(* IEC 61131-3 sources: 2026_Projet_YGO_ExcavatriceDragage/TOOLS/TEST_AUTO_CI/RESULTS/H_TREUILS_BENNE/tests (part 4) *)

(* ---- test_fb_winchoutputinterlock.st ---- *)
(* =======================================================================
   🧪 test_fb_winchoutputinterlock.st — FB_WinchOutputInterlock (TC-P10-012, 013, 020, 021, 022, 039.1)
   ───────────────────────────────────────────────────────────────
   Fiche : DOC/AF/AF_Partie-10_Fonction_Winch/FB_WinchOutputInterlock_v1.0.md
   Conventions : 1 appel fb() = 1 scan ; ADVANCE_TIME(10000000) entre les
   scans pour les fronts R_TRIG ; hex décrit en décimal (bit 0 = 1).
   Watchdog frein = 500ms ; RestartDelay = 1500ms ; DeadTimeSameDir/OppositeDir = 1s (défaut).
   Maintien §3bis : DropConfirmDelay = 100ms , MaxSenseHoldTime (T_max) = 1s (défauts, AC8).
   ======================================================================= *)

SETUP
VAR
    fb : FB_WinchOutputInterlock;
END_VAR
END_SETUP

(* ── Remise à zéro commune : Enable=TRUE, frein serré, pause 1500ms pour purger RestartRequired/DeadTime ── *)

TEST 'TC-P10-012 Watchdog frein : BrakeCmd sans confirmation 500ms -> bit0, RestartInhibit, FAULT ; pas de faux defaut au RestartRequired'
    (* Scan 1 : regime nominal, frein serre (BrakeFeedback=FALSE), pause pour purger *)
    fb(Enable := TRUE, Reset := FALSE, SafeStop := FALSE, AscentPermit := TRUE, DescendPermit := TRUE, PowerContactorEngaged := TRUE,
       BrakeFeedback := FALSE, FwdRevSpeedFeedbackOff := TRUE,
       RequestedRelayFwd := FALSE, RequestedRelayRev := FALSE,
       RequestedContactor1 := FALSE, RequestedContactor2 := FALSE,
       RequestedContactor3 := FALSE, RequestedContactor4 := FALSE,
       RequestedStep := 0);
    ADVANCE_TIME(1500000000);
fb(Enable := TRUE, Reset := FALSE, SafeStop := FALSE, AscentPermit := TRUE, DescendPermit := TRUE, PowerContactorEngaged := TRUE,
       BrakeFeedback := FALSE, FwdRevSpeedFeedbackOff := TRUE,
       RequestedRelayFwd := FALSE, RequestedRelayRev := FALSE,
       RequestedContactor1 := FALSE, RequestedContactor2 := FALSE,
       RequestedContactor3 := FALSE, RequestedContactor4 := FALSE,
       RequestedStep := 0);
    ASSERT_TRUE(fb.Ready, 'Regime nominal -> Ready=TRUE');

    (* Scan 2 : demande mouvement, frein NON confirme ouvert (BrakeFeedback=FALSE) -> watchdog arme *)
    ADVANCE_TIME(10000000);
fb(Enable := TRUE, Reset := FALSE, SafeStop := FALSE, AscentPermit := TRUE, DescendPermit := TRUE, PowerContactorEngaged := TRUE,
       BrakeFeedback := FALSE, FwdRevSpeedFeedbackOff := TRUE,
       RequestedRelayFwd := TRUE, RequestedRelayRev := FALSE,
       RequestedContactor1 := TRUE, RequestedContactor2 := FALSE,
       RequestedContactor3 := FALSE, RequestedContactor4 := FALSE,
       RequestedStep := 1);
    ASSERT_TRUE(fb.RelayFwd, 'Demande montee -> RelayFwd');
    ASSERT_TRUE(fb.BrakeCmd, 'Demande montee -> BrakeCmd');
    ASSERT_EQ(fb.State, E_WinchFinalInterlockState.WAIT_BRAKE_COMMAND_CONFIRMATION, 'Etat WAIT_BRAKE_COMMAND_CONFIRMATION (2)');

    (* Scan 3 : apres 500ms sans confirmation -> defaut frein *)
    ADVANCE_TIME(500000000);
fb(Enable := TRUE, Reset := FALSE, SafeStop := FALSE, AscentPermit := TRUE, DescendPermit := TRUE, PowerContactorEngaged := TRUE,
       BrakeFeedback := FALSE, FwdRevSpeedFeedbackOff := TRUE,
       RequestedRelayFwd := TRUE, RequestedRelayRev := FALSE,
       RequestedContactor1 := TRUE, RequestedContactor2 := FALSE,
       RequestedContactor3 := FALSE, RequestedContactor4 := FALSE,
       RequestedStep := 1);
    ASSERT_TRUE(fb.Error, 'Timeout frein 500ms -> Error');
    ASSERT_EQ(fb.ErrorId, 1, 'Timeout frein -> bit0 (1)');
    ASSERT_TRUE(fb.RestartInhibit, 'Timeout frein -> RestartInhibit=TRUE');
    ASSERT_EQ(fb.Reason, E_WinchFinalInterlockReason.BRAKE_COMMAND_NOT_CONFIRMED, 'Reason=BRAKE_COMMAND_NOT_CONFIRMED (1)');
    ASSERT_EQ(fb.State, E_WinchFinalInterlockState.FAULT, 'Etat FAULT (5)');
END_TEST

TEST 'TC-P10-012bis Pas de faux defaut au RestartRequired : BrakeCmd retenu ne doit pas armer le watchdog'
    (* Scan 1 : regime nominal, pause pour purger *)
    fb(Enable := TRUE, Reset := FALSE, SafeStop := FALSE, AscentPermit := TRUE, DescendPermit := TRUE, PowerContactorEngaged := TRUE,
       BrakeFeedback := FALSE, FwdRevSpeedFeedbackOff := TRUE,
       RequestedRelayFwd := FALSE, RequestedRelayRev := FALSE,
       RequestedContactor1 := FALSE, RequestedContactor2 := FALSE,
       RequestedContactor3 := FALSE, RequestedContactor4 := FALSE,
       RequestedStep := 0);
    ADVANCE_TIME(1500000000);
fb(Enable := TRUE, Reset := FALSE, SafeStop := FALSE, AscentPermit := TRUE, DescendPermit := TRUE, PowerContactorEngaged := TRUE,
       BrakeFeedback := FALSE, FwdRevSpeedFeedbackOff := TRUE,
       RequestedRelayFwd := FALSE, RequestedRelayRev := FALSE,
       RequestedContactor1 := FALSE, RequestedContactor2 := FALSE,
       RequestedContactor3 := FALSE, RequestedContactor4 := FALSE,
       RequestedStep := 0);

    (* Scan 2 : demande mouvement, frein confirme (BrakeFeedback=TRUE) -> mouvement autorise *)
    ADVANCE_TIME(10000000);
fb(Enable := TRUE, Reset := FALSE, SafeStop := FALSE, AscentPermit := TRUE, DescendPermit := TRUE, PowerContactorEngaged := TRUE,
       BrakeFeedback := TRUE, FwdRevSpeedFeedbackOff := TRUE,
       RequestedRelayFwd := TRUE, RequestedRelayRev := FALSE,
       RequestedContactor1 := TRUE, RequestedContactor2 := FALSE,
       RequestedContactor3 := FALSE, RequestedContactor4 := FALSE,
       RequestedStep := 1);
    ASSERT_TRUE(fb.RelayFwd, 'Mouvement autorise -> RelayFwd');

    (* Scan 3 : arret -> RestartRequired=TRUE *)
    ADVANCE_TIME(10000000);
fb(Enable := TRUE, Reset := FALSE, SafeStop := FALSE, AscentPermit := TRUE, DescendPermit := TRUE, PowerContactorEngaged := TRUE,
       BrakeFeedback := FALSE, FwdRevSpeedFeedbackOff := TRUE,
       RequestedRelayFwd := FALSE, RequestedRelayRev := FALSE,
       RequestedContactor1 := FALSE, RequestedContactor2 := FALSE,
       RequestedContactor3 := FALSE, RequestedContactor4 := FALSE,
       RequestedStep := 0);

    (* Scan 4 : nouvelle demande IMMEDIATE (RestartRequired=TRUE) -> BrakeCmd retenu, watchdog NON arme *)
    ADVANCE_TIME(10000000);
fb(Enable := TRUE, Reset := FALSE, SafeStop := FALSE, AscentPermit := TRUE, DescendPermit := TRUE, PowerContactorEngaged := TRUE,
       BrakeFeedback := FALSE, FwdRevSpeedFeedbackOff := TRUE,
       RequestedRelayFwd := TRUE, RequestedRelayRev := FALSE,
       RequestedContactor1 := TRUE, RequestedContactor2 := FALSE,
       RequestedContactor3 := FALSE, RequestedContactor4 := FALSE,
       RequestedStep := 1);
    ASSERT_FALSE(fb.RelayFwd, 'RestartRequired -> RelayFwd retenu');
    ASSERT_FALSE(fb.BrakeCmd, 'RestartRequired -> BrakeCmd retenu (FALSE)');
    ASSERT_EQ(fb.State, E_WinchFinalInterlockState.WAIT_RESTART_DELAY, 'Etat WAIT_RESTART_DELAY (4)');

    (* Scan 5 : apres 500ms, BrakeCmd=FALSE -> PAS de faux defaut *)
    ADVANCE_TIME(500000000);
fb(Enable := TRUE, Reset := FALSE, SafeStop := FALSE, AscentPermit := TRUE, DescendPermit := TRUE, PowerContactorEngaged := TRUE,
       BrakeFeedback := FALSE, FwdRevSpeedFeedbackOff := TRUE,
       RequestedRelayFwd := TRUE, RequestedRelayRev := FALSE,
       RequestedContactor1 := TRUE, RequestedContactor2 := FALSE,
       RequestedContactor3 := FALSE, RequestedContactor4 := FALSE,
       RequestedStep := 1);
    ASSERT_FALSE(fb.Error, 'BrakeCmd retenu par RestartRequired -> PAS de faux defaut frein');
    ASSERT_FALSE(fb.RestartInhibit, 'Pas de RestartInhibit sur faux defaut');
END_TEST

TEST 'TC-P10-013 Defaut frein : latches preserves hors Enable, reautorisation complete'
    (* Scan 1 : regime nominal, pause pour purger *)
    fb(Enable := TRUE, Reset := FALSE, SafeStop := FALSE, AscentPermit := TRUE, DescendPermit := TRUE, PowerContactorEngaged := TRUE,
       BrakeFeedback := FALSE, FwdRevSpeedFeedbackOff := TRUE,
       RequestedRelayFwd := FALSE, RequestedRelayRev := FALSE,
       RequestedContactor1 := FALSE, RequestedContactor2 := FALSE,
       RequestedContactor3 := FALSE, RequestedContactor4 := FALSE,
       RequestedStep := 0);
    ADVANCE_TIME(1500000000);
fb(Enable := TRUE, Reset := FALSE, SafeStop := FALSE, AscentPermit := TRUE, DescendPermit := TRUE, PowerContactorEngaged := TRUE,
       BrakeFeedback := FALSE, FwdRevSpeedFeedbackOff := TRUE,
       RequestedRelayFwd := FALSE, RequestedRelayRev := FALSE,
       RequestedContactor1 := FALSE, RequestedContactor2 := FALSE,
       RequestedContactor3 := FALSE, RequestedContactor4 := FALSE,
       RequestedStep := 0);

    (* Scan 2 : demande mouvement, frein non confirme -> watchdog arme *)
    ADVANCE_TIME(10000000);
fb(Enable := TRUE, Reset := FALSE, SafeStop := FALSE, AscentPermit := TRUE, DescendPermit := TRUE, PowerContactorEngaged := TRUE,
       BrakeFeedback := FALSE, FwdRevSpeedFeedbackOff := TRUE,
       RequestedRelayFwd := TRUE, RequestedRelayRev := FALSE,
       RequestedContactor1 := TRUE, RequestedContactor2 := FALSE,
       RequestedContactor3 := FALSE, RequestedContactor4 := FALSE,
       RequestedStep := 1);
    ADVANCE_TIME(500000000);
fb(Enable := TRUE, Reset := FALSE, SafeStop := FALSE, AscentPermit := TRUE, DescendPermit := TRUE, PowerContactorEngaged := TRUE,
       BrakeFeedback := FALSE, FwdRevSpeedFeedbackOff := TRUE,
       RequestedRelayFwd := TRUE, RequestedRelayRev := FALSE,
       RequestedContactor1 := TRUE, RequestedContactor2 := FALSE,
       RequestedContactor3 := FALSE, RequestedContactor4 := FALSE,
       RequestedStep := 1);
    ASSERT_TRUE(fb.Error, 'Precondition : defaut frein');
    ASSERT_TRUE(fb.RestartInhibit, 'Precondition : RestartInhibit');

    (* Scan 3 : Enable=FALSE -> sorties FALSE MAIS latches preserves *)
    ADVANCE_TIME(10000000);
    fb(Enable := FALSE, Reset := FALSE, SafeStop := FALSE, PowerContactorEngaged := TRUE,
       BrakeFeedback := FALSE, FwdRevSpeedFeedbackOff := TRUE,
       RequestedRelayFwd := TRUE, RequestedRelayRev := FALSE,
       RequestedContactor1 := TRUE, RequestedContactor2 := FALSE,
       RequestedContactor3 := FALSE, RequestedContactor4 := FALSE,
       RequestedStep := 1);
    ASSERT_FALSE(fb.RelayFwd, 'Enable=FALSE -> RelayFwd=FALSE');
    ASSERT_FALSE(fb.BrakeCmd, 'Enable=FALSE -> BrakeCmd=FALSE');
    ASSERT_TRUE(fb.RestartInhibit, 'Enable=FALSE -> RestartInhibit PRESERVE');
    ASSERT_EQ(fb.ErrorId, 1, 'Enable=FALSE -> ErrorId bit0 PRESERVE');

    (* Scan 4 : re-Enable, cause disparue (BrakeFeedback=TRUE) + front Reset -> ResetRequired leve *)
    ADVANCE_TIME(10000000);
    fb(Enable := TRUE, Reset := TRUE, SafeStop := FALSE, PowerContactorEngaged := TRUE,
       BrakeFeedback := TRUE, FwdRevSpeedFeedbackOff := TRUE,
       RequestedRelayFwd := FALSE, RequestedRelayRev := FALSE,
       RequestedContactor1 := FALSE, RequestedContactor2 := FALSE,
       RequestedContactor3 := FALSE, RequestedContactor4 := FALSE,
       RequestedStep := 0);
    ADVANCE_TIME(10000000);
fb(Enable := TRUE, Reset := FALSE, SafeStop := FALSE, AscentPermit := TRUE, DescendPermit := TRUE, PowerContactorEngaged := TRUE,
       BrakeFeedback := TRUE, FwdRevSpeedFeedbackOff := TRUE,
       RequestedRelayFwd := FALSE, RequestedRelayRev := FALSE,
       RequestedContactor1 := FALSE, RequestedContactor2 := FALSE,
       RequestedContactor3 := FALSE, RequestedContactor4 := FALSE,
       RequestedStep := 0);
    ASSERT_FALSE(fb.Error, 'Cause disparue + Reset -> Error=FALSE');

    (* Scan 5 : demande neutre observee (MotorRequest=FALSE) -> NeutralRequestSeen *)
    ADVANCE_TIME(10000000);
fb(Enable := TRUE, Reset := FALSE, SafeStop := FALSE, AscentPermit := TRUE, DescendPermit := TRUE, PowerContactorEngaged := TRUE,
       BrakeFeedback := FALSE, FwdRevSpeedFeedbackOff := TRUE,
       RequestedRelayFwd := FALSE, RequestedRelayRev := FALSE,
       RequestedContactor1 := FALSE, RequestedContactor2 := FALSE,
       RequestedContactor3 := FALSE, RequestedContactor4 := FALSE,
       RequestedStep := 0);
    ADVANCE_TIME(1500000000);
fb(Enable := TRUE, Reset := FALSE, SafeStop := FALSE, AscentPermit := TRUE, DescendPermit := TRUE, PowerContactorEngaged := TRUE,
       BrakeFeedback := FALSE, FwdRevSpeedFeedbackOff := TRUE,
       RequestedRelayFwd := FALSE, RequestedRelayRev := FALSE,
       RequestedContactor1 := FALSE, RequestedContactor2 := FALSE,
       RequestedContactor3 := FALSE, RequestedContactor4 := FALSE,
       RequestedStep := 0);

    (* Scan 6 : nouvelle demande distincte -> RestartInhibit leve *)
    ADVANCE_TIME(10000000);
fb(Enable := TRUE, Reset := FALSE, SafeStop := FALSE, AscentPermit := TRUE, DescendPermit := TRUE, PowerContactorEngaged := TRUE,
       BrakeFeedback := TRUE, FwdRevSpeedFeedbackOff := TRUE,
       RequestedRelayFwd := TRUE, RequestedRelayRev := FALSE,
       RequestedContactor1 := TRUE, RequestedContactor2 := FALSE,
       RequestedContactor3 := FALSE, RequestedContactor4 := FALSE,
       RequestedStep := 1);
    ASSERT_FALSE(fb.RestartInhibit, 'Reautorisation complete -> RestartInhibit=FALSE');
    ASSERT_TRUE(fb.RelayFwd, 'Reautorisation -> mouvement autorise');
END_TEST

TEST 'TC-P10-020 Watchdog frein reel terrain : temps/contacteur/bobine'
    (* (essai site — stub) : le watchdog frein reel (temps de reponse contacteur/bobine, usure)
       est une verification terrain sur l automate reel, jamais automatisable en boite noire.
       On verifie ici la brique logicielle : le watchdog 500ms se declenche sur BrakeCmd sans
       confirmation, condition necessaire du diagnostic terrain. *)
    fb(Enable := TRUE, Reset := FALSE, SafeStop := FALSE, AscentPermit := TRUE, DescendPermit := TRUE, PowerContactorEngaged := TRUE,
       BrakeFeedback := FALSE, FwdRevSpeedFeedbackOff := TRUE,
       RequestedRelayFwd := FALSE, RequestedRelayRev := FALSE,
       RequestedContactor1 := FALSE, RequestedContactor2 := FALSE,
       RequestedContactor3 := FALSE, RequestedContactor4 := FALSE,
       RequestedStep := 0);
    ADVANCE_TIME(1500000000);
    // Scan neutre temporise : purge RestartRequired/DeadTimePending (TON tickes apres la pause,
    // comme les ~150 scans de 10ms d'une vraie pause automate) avant la demande mouvement.
fb(Enable := TRUE, Reset := FALSE, SafeStop := FALSE, AscentPermit := TRUE, DescendPermit := TRUE, PowerContactorEngaged := TRUE,
       BrakeFeedback := FALSE, FwdRevSpeedFeedbackOff := TRUE,
       RequestedRelayFwd := FALSE, RequestedRelayRev := FALSE,
       RequestedContactor1 := FALSE, RequestedContactor2 := FALSE,
       RequestedContactor3 := FALSE, RequestedContactor4 := FALSE,
       RequestedStep := 0);
    ADVANCE_TIME(10000000);
fb(Enable := TRUE, Reset := FALSE, SafeStop := FALSE, AscentPermit := TRUE, DescendPermit := TRUE, PowerContactorEngaged := TRUE,
       BrakeFeedback := FALSE, FwdRevSpeedFeedbackOff := TRUE,
       RequestedRelayFwd := TRUE, RequestedRelayRev := FALSE,
       RequestedContactor1 := TRUE, RequestedContactor2 := FALSE,
       RequestedContactor3 := FALSE, RequestedContactor4 := FALSE,
       RequestedStep := 1);
    ADVANCE_TIME(500000000);
fb(Enable := TRUE, Reset := FALSE, SafeStop := FALSE, AscentPermit := TRUE, DescendPermit := TRUE, PowerContactorEngaged := TRUE,
       BrakeFeedback := FALSE, FwdRevSpeedFeedbackOff := TRUE,
       RequestedRelayFwd := TRUE, RequestedRelayRev := FALSE,
       RequestedContactor1 := TRUE, RequestedContactor2 := FALSE,
       RequestedContactor3 := FALSE, RequestedContactor4 := FALSE,
       RequestedStep := 1);
    ASSERT_TRUE(fb.Error, 'Watchdog frein logiciel 500ms -> Error (brique du diagnostic terrain)');
    ASSERT_EQ(fb.Reason, E_WinchFinalInterlockReason.BRAKE_COMMAND_NOT_CONFIRMED, 'Reason=BRAKE_COMMAND_NOT_CONFIRMED');
END_TEST

TEST 'TC-P10-021 Temps mort meme sens : 1s apres arret -> nouvelle demande (DeadTimeSameDir)'
    (* DeadTimeSameDir=2s force pour rendre le temps mort observable (par defaut 1s, masque
       par RestartDelay 1500ms). La demande meme sens est retenue tant que DeadTimeSameDir
       n est pas ecoule. *)
    fb(Enable := TRUE, Reset := FALSE, SafeStop := FALSE, AscentPermit := TRUE, DescendPermit := TRUE, PowerContactorEngaged := TRUE,
       BrakeFeedback := FALSE, FwdRevSpeedFeedbackOff := TRUE,
       RequestedRelayFwd := FALSE, RequestedRelayRev := FALSE,
       RequestedContactor1 := FALSE, RequestedContactor2 := FALSE,
       RequestedContactor3 := FALSE, RequestedContactor4 := FALSE,
       RequestedStep := 0, DeadTimeSameDir := T#2s, DeadTimeOppositeDir := T#2s);
    ADVANCE_TIME(1500000000);
fb(Enable := TRUE, Reset := FALSE, SafeStop := FALSE, AscentPermit := TRUE, DescendPermit := TRUE, PowerContactorEngaged := TRUE,
       BrakeFeedback := FALSE, FwdRevSpeedFeedbackOff := TRUE,
       RequestedRelayFwd := FALSE, RequestedRelayRev := FALSE,
       RequestedContactor1 := FALSE, RequestedContactor2 := FALSE,
       RequestedContactor3 := FALSE, RequestedContactor4 := FALSE,
       RequestedStep := 0, DeadTimeSameDir := T#2s, DeadTimeOppositeDir := T#2s);

    (* Scan 2 : demande montee, frein confirme -> mouvement *)
    ADVANCE_TIME(10000000);
fb(Enable := TRUE, Reset := FALSE, SafeStop := FALSE, AscentPermit := TRUE, DescendPermit := TRUE, PowerContactorEngaged := TRUE,
       BrakeFeedback := TRUE, FwdRevSpeedFeedbackOff := TRUE,
       RequestedRelayFwd := TRUE, RequestedRelayRev := FALSE,
       RequestedContactor1 := TRUE, RequestedContactor2 := FALSE,
       RequestedContactor3 := FALSE, RequestedContactor4 := FALSE,
       RequestedStep := 1, DeadTimeSameDir := T#2s, DeadTimeOppositeDir := T#2s);
    ASSERT_TRUE(fb.RelayFwd, 'Mouvement autorise -> RelayFwd');

    (* Scan 3 : arret -> DeadTimePending=TRUE *)
    ADVANCE_TIME(10000000);
fb(Enable := TRUE, Reset := FALSE, SafeStop := FALSE, AscentPermit := TRUE, DescendPermit := TRUE, PowerContactorEngaged := TRUE,
       BrakeFeedback := FALSE, FwdRevSpeedFeedbackOff := TRUE,
       RequestedRelayFwd := FALSE, RequestedRelayRev := FALSE,
       RequestedContactor1 := FALSE, RequestedContactor2 := FALSE,
       RequestedContactor3 := FALSE, RequestedContactor4 := FALSE,
       RequestedStep := 0, DeadTimeSameDir := T#2s, DeadTimeOppositeDir := T#2s);

    (* Scan 4 : apres 1500ms (RestartRequired leve), DeadTimeSameDir=2s pas encore ecoule -> retenu *)
    ADVANCE_TIME(1500000000);
fb(Enable := TRUE, Reset := FALSE, SafeStop := FALSE, AscentPermit := TRUE, DescendPermit := TRUE, PowerContactorEngaged := TRUE,
       BrakeFeedback := FALSE, FwdRevSpeedFeedbackOff := TRUE,
       RequestedRelayFwd := TRUE, RequestedRelayRev := FALSE,
       RequestedContactor1 := TRUE, RequestedContactor2 := FALSE,
       RequestedContactor3 := FALSE, RequestedContactor4 := FALSE,
       RequestedStep := 1, DeadTimeSameDir := T#2s, DeadTimeOppositeDir := T#2s);
    ASSERT_FALSE(fb.RelayFwd, 'DeadTimeSameDir pas ecoule -> demande meme sens retenue');
    ASSERT_EQ(fb.State, E_WinchFinalInterlockState.WAIT_RESTART_DELAY, 'Etat WAIT_RESTART_DELAY (4)');

    (* Scan 5 : apres 2s (DeadTimeSameDir ecoule) -> demande meme sens acceptee *)
    ADVANCE_TIME(600000000);
fb(Enable := TRUE, Reset := FALSE, SafeStop := FALSE, AscentPermit := TRUE, DescendPermit := TRUE, PowerContactorEngaged := TRUE,
       BrakeFeedback := TRUE, FwdRevSpeedFeedbackOff := TRUE,
       RequestedRelayFwd := TRUE, RequestedRelayRev := FALSE,
       RequestedContactor1 := TRUE, RequestedContactor2 := FALSE,
       RequestedContactor3 := FALSE, RequestedContactor4 := FALSE,
       RequestedStep := 1, DeadTimeSameDir := T#2s, DeadTimeOppositeDir := T#2s);
    ASSERT_TRUE(fb.RelayFwd, 'DeadTimeSameDir ecoule -> demande meme sens acceptee');
END_TEST

TEST 'TC-P10-022 Temps mort inversion : 1s apres arret + inversion sens (DeadTimeOppositeDir)'
    (* DeadTimeOppositeDir=2s force pour rendre le temps mort d inversion observable.
       L inversion est retenue tant que DeadTimeOppositeDir n est pas ecoule. *)
    fb(Enable := TRUE, Reset := FALSE, SafeStop := FALSE, AscentPermit := TRUE, DescendPermit := TRUE, PowerContactorEngaged := TRUE,
       BrakeFeedback := FALSE, FwdRevSpeedFeedbackOff := TRUE,
       RequestedRelayFwd := FALSE, RequestedRelayRev := FALSE,
       RequestedContactor1 := FALSE, RequestedContactor2 := FALSE,
       RequestedContactor3 := FALSE, RequestedContactor4 := FALSE,
       RequestedStep := 0, DeadTimeSameDir := T#1s, DeadTimeOppositeDir := T#2s);
    ADVANCE_TIME(1500000000);
fb(Enable := TRUE, Reset := FALSE, SafeStop := FALSE, AscentPermit := TRUE, DescendPermit := TRUE, PowerContactorEngaged := TRUE,
       BrakeFeedback := FALSE, FwdRevSpeedFeedbackOff := TRUE,
       RequestedRelayFwd := FALSE, RequestedRelayRev := FALSE,
       RequestedContactor1 := FALSE, RequestedContactor2 := FALSE,
       RequestedContactor3 := FALSE, RequestedContactor4 := FALSE,
       RequestedStep := 0, DeadTimeSameDir := T#1s, DeadTimeOppositeDir := T#2s);

    (* Scan 2 : demande montee, frein confirme -> mouvement *)
    ADVANCE_TIME(10000000);
fb(Enable := TRUE, Reset := FALSE, SafeStop := FALSE, AscentPermit := TRUE, DescendPermit := TRUE, PowerContactorEngaged := TRUE,
       BrakeFeedback := TRUE, FwdRevSpeedFeedbackOff := TRUE,
       RequestedRelayFwd := TRUE, RequestedRelayRev := FALSE,
       RequestedContactor1 := TRUE, RequestedContactor2 := FALSE,
       RequestedContactor3 := FALSE, RequestedContactor4 := FALSE,
       RequestedStep := 1, DeadTimeSameDir := T#1s, DeadTimeOppositeDir := T#2s);
    ASSERT_TRUE(fb.RelayFwd, 'Mouvement montee -> RelayFwd');

    (* Scan 3 : arret -> DeadTimePending=TRUE *)
    ADVANCE_TIME(10000000);
fb(Enable := TRUE, Reset := FALSE, SafeStop := FALSE, AscentPermit := TRUE, DescendPermit := TRUE, PowerContactorEngaged := TRUE,
       BrakeFeedback := FALSE, FwdRevSpeedFeedbackOff := TRUE,
       RequestedRelayFwd := FALSE, RequestedRelayRev := FALSE,
       RequestedContactor1 := FALSE, RequestedContactor2 := FALSE,
       RequestedContactor3 := FALSE, RequestedContactor4 := FALSE,
       RequestedStep := 0, DeadTimeSameDir := T#1s, DeadTimeOppositeDir := T#2s);

    (* Scan 4 : apres 1500ms, inversion (descente) -> DeadTimeOppositeDir=2s pas ecoule -> retenu *)
    ADVANCE_TIME(1500000000);
fb(Enable := TRUE, Reset := FALSE, SafeStop := FALSE, AscentPermit := TRUE, DescendPermit := TRUE, PowerContactorEngaged := TRUE,
       BrakeFeedback := FALSE, FwdRevSpeedFeedbackOff := TRUE,
       RequestedRelayFwd := FALSE, RequestedRelayRev := TRUE,
       RequestedContactor1 := TRUE, RequestedContactor2 := FALSE,
       RequestedContactor3 := FALSE, RequestedContactor4 := FALSE,
       RequestedStep := 1, DeadTimeSameDir := T#1s, DeadTimeOppositeDir := T#2s);
    ASSERT_FALSE(fb.RelayRev, 'DeadTimeOppositeDir pas ecoule -> inversion retenue');
    ASSERT_EQ(fb.State, E_WinchFinalInterlockState.WAIT_RESTART_DELAY, 'Etat WAIT_RESTART_DELAY (4)');

    (* Scan 5 : apres 2s (DeadTimeOppositeDir ecoule) -> inversion acceptee *)
    ADVANCE_TIME(600000000);
fb(Enable := TRUE, Reset := FALSE, SafeStop := FALSE, AscentPermit := TRUE, DescendPermit := TRUE, PowerContactorEngaged := TRUE,
       BrakeFeedback := TRUE, FwdRevSpeedFeedbackOff := TRUE,
       RequestedRelayFwd := FALSE, RequestedRelayRev := TRUE,
       RequestedContactor1 := TRUE, RequestedContactor2 := FALSE,
       RequestedContactor3 := FALSE, RequestedContactor4 := FALSE,
       RequestedStep := 1, DeadTimeSameDir := T#1s, DeadTimeOppositeDir := T#2s);
    ASSERT_TRUE(fb.RelayRev, 'DeadTimeOppositeDir ecoule -> inversion acceptee');
END_TEST

TEST 'TC-P10-039.1 Frein couple direct : BrakeCmd = RelayFwd OR RelayRev dans tous les etats'
    (* Scan 1 : regime nominal, pause pour purger *)
    fb(Enable := TRUE, Reset := FALSE, SafeStop := FALSE, AscentPermit := TRUE, DescendPermit := TRUE, PowerContactorEngaged := TRUE,
       BrakeFeedback := FALSE, FwdRevSpeedFeedbackOff := TRUE,
       RequestedRelayFwd := FALSE, RequestedRelayRev := FALSE,
       RequestedContactor1 := FALSE, RequestedContactor2 := FALSE,
       RequestedContactor3 := FALSE, RequestedContactor4 := FALSE,
       RequestedStep := 0);
    ADVANCE_TIME(1500000000);
fb(Enable := TRUE, Reset := FALSE, SafeStop := FALSE, AscentPermit := TRUE, DescendPermit := TRUE, PowerContactorEngaged := TRUE,
       BrakeFeedback := FALSE, FwdRevSpeedFeedbackOff := TRUE,
       RequestedRelayFwd := FALSE, RequestedRelayRev := FALSE,
       RequestedContactor1 := FALSE, RequestedContactor2 := FALSE,
       RequestedContactor3 := FALSE, RequestedContactor4 := FALSE,
       RequestedStep := 0);
    ASSERT_FALSE(fb.BrakeCmd, 'Repos : BrakeCmd=FALSE (RelayFwd/Rev=FALSE)');

    (* Scan 2 : mouvement montee -> BrakeCmd=TRUE (RelayFwd=TRUE) *)
    ADVANCE_TIME(10000000);
fb(Enable := TRUE, Reset := FALSE, SafeStop := FALSE, AscentPermit := TRUE, DescendPermit := TRUE, PowerContactorEngaged := TRUE,
       BrakeFeedback := TRUE, FwdRevSpeedFeedbackOff := TRUE,
       RequestedRelayFwd := TRUE, RequestedRelayRev := FALSE,
       RequestedContactor1 := TRUE, RequestedContactor2 := FALSE,
       RequestedContactor3 := FALSE, RequestedContactor4 := FALSE,
       RequestedStep := 1);
    ASSERT_TRUE(fb.RelayFwd, 'Mouvement -> RelayFwd=TRUE');
    ASSERT_TRUE(fb.BrakeCmd, 'Mouvement -> BrakeCmd=TRUE (couple direct)');

    (* Scan 3 : arret -> BrakeCmd=FALSE *)
    ADVANCE_TIME(10000000);
fb(Enable := TRUE, Reset := FALSE, SafeStop := FALSE, AscentPermit := TRUE, DescendPermit := TRUE, PowerContactorEngaged := TRUE,
       BrakeFeedback := FALSE, FwdRevSpeedFeedbackOff := TRUE,
       RequestedRelayFwd := FALSE, RequestedRelayRev := FALSE,
       RequestedContactor1 := FALSE, RequestedContactor2 := FALSE,
       RequestedContactor3 := FALSE, RequestedContactor4 := FALSE,
       RequestedStep := 0);
    ASSERT_FALSE(fb.RelayFwd, 'Arret -> RelayFwd=FALSE');
    ASSERT_FALSE(fb.BrakeCmd, 'Arret -> BrakeCmd=FALSE (jamais de divergence frein/mouvement)');
END_TEST

TEST 'TC-P10-023a §3bis : sens maintenu apres chute de palier a 0 tant que contacteurs non confirmes, puis chute sur DropConfirmDelay'
    (* Chute de palier : RequestedStep -> 0 mais RequestedRelayFwd reste TRUE (demande transitoire
       FB_Winch). La barriere TIENT le contacteur de sens jusqu a FwdRevSpeedFeedbackOff confirme
       (debounced DropConfirmDelay=300ms) OU T_max. Aucun faux arret pendant le debounce. *)
    fb(Enable := TRUE, Reset := FALSE, SafeStop := FALSE, AscentPermit := TRUE, DescendPermit := TRUE, PowerContactorEngaged := TRUE,
       BrakeFeedback := FALSE, FwdRevSpeedFeedbackOff := TRUE,
       RequestedRelayFwd := FALSE, RequestedRelayRev := FALSE,
       RequestedContactor1 := FALSE, RequestedContactor2 := FALSE,
       RequestedContactor3 := FALSE, RequestedContactor4 := FALSE,
       RequestedStep := 0, DropConfirmDelay := T#300ms, MaxSenseHoldTime := T#1s);
    ADVANCE_TIME(1500000000);
fb(Enable := TRUE, Reset := FALSE, SafeStop := FALSE, AscentPermit := TRUE, DescendPermit := TRUE, PowerContactorEngaged := TRUE,
       BrakeFeedback := FALSE, FwdRevSpeedFeedbackOff := TRUE,
       RequestedRelayFwd := FALSE, RequestedRelayRev := FALSE,
       RequestedContactor1 := FALSE, RequestedContactor2 := FALSE,
       RequestedContactor3 := FALSE, RequestedContactor4 := FALSE,
       RequestedStep := 0, DropConfirmDelay := T#300ms, MaxSenseHoldTime := T#1s);
    ASSERT_TRUE(fb.Ready, 'Regime nominal -> Ready=TRUE');

    (* Scan 2 : mouvement montee, frein confirme, contacteurs engages (FwdRevSpeedFeedbackOff=FALSE) *)
    ADVANCE_TIME(10000000);
fb(Enable := TRUE, Reset := FALSE, SafeStop := FALSE, AscentPermit := TRUE, DescendPermit := TRUE, PowerContactorEngaged := TRUE,
       BrakeFeedback := TRUE, FwdRevSpeedFeedbackOff := FALSE,
       RequestedRelayFwd := TRUE, RequestedRelayRev := FALSE,
       RequestedContactor1 := TRUE, RequestedContactor2 := FALSE,
       RequestedContactor3 := FALSE, RequestedContactor4 := FALSE,
       RequestedStep := 1, DropConfirmDelay := T#300ms, MaxSenseHoldTime := T#1s);
    ASSERT_TRUE(fb.RelayFwd, 'Mouvement -> RelayFwd');
    ASSERT_TRUE(fb.BrakeCmd, 'Mouvement -> BrakeCmd');

    (* Scan 3 : chute a palier 0, RequestedRelayFwd TOUJOURS TRUE, contacteurs pas encore retombes *)
    ADVANCE_TIME(10000000);
fb(Enable := TRUE, Reset := FALSE, SafeStop := FALSE, AscentPermit := TRUE, DescendPermit := TRUE, PowerContactorEngaged := TRUE,
       BrakeFeedback := TRUE, FwdRevSpeedFeedbackOff := FALSE,
       RequestedRelayFwd := TRUE, RequestedRelayRev := FALSE,
       RequestedContactor1 := FALSE, RequestedContactor2 := FALSE,
       RequestedContactor3 := FALSE, RequestedContactor4 := FALSE,
       RequestedStep := 0, DropConfirmDelay := T#300ms, MaxSenseHoldTime := T#1s);
    ASSERT_TRUE(fb.RelayFwd, 'Chute palier -> contacteur de sens MAINTENU (§3bis)');
    ASSERT_TRUE(fb.BrakeCmd, 'Maintien -> BrakeCmd reste TRUE (couple direct)');
    ASSERT_TRUE(fb.SenseHoldActive, 'Diag SenseHoldActive');
    ASSERT_EQ(fb.State, E_WinchFinalInterlockState.WAIT_SENSE_DROP_CONFIRM, 'Etat WAIT_SENSE_DROP_CONFIRM (6)');

    (* Scan 4 : feedback retombee percu (FwdRevSpeedFeedbackOff=TRUE) mais debounce pas ecoule -> tenu *)
    ADVANCE_TIME(100000000);
fb(Enable := TRUE, Reset := FALSE, SafeStop := FALSE, AscentPermit := TRUE, DescendPermit := TRUE, PowerContactorEngaged := TRUE,
       BrakeFeedback := TRUE, FwdRevSpeedFeedbackOff := TRUE,
       RequestedRelayFwd := TRUE, RequestedRelayRev := FALSE,
       RequestedContactor1 := FALSE, RequestedContactor2 := FALSE,
       RequestedContactor3 := FALSE, RequestedContactor4 := FALSE,
       RequestedStep := 0, DropConfirmDelay := T#300ms, MaxSenseHoldTime := T#1s);
    ASSERT_TRUE(fb.RelayFwd, 'Debounce DropConfirmDelay pas ecoule -> sens TOUJOURS tenu (AC7)');

    (* Scan 5 : DropConfirmDelay (300ms) ecoule -> chute normale du sens *)
    ADVANCE_TIME(300000000);
fb(Enable := TRUE, Reset := FALSE, SafeStop := FALSE, AscentPermit := TRUE, DescendPermit := TRUE, PowerContactorEngaged := TRUE,
       BrakeFeedback := TRUE, FwdRevSpeedFeedbackOff := TRUE,
       RequestedRelayFwd := TRUE, RequestedRelayRev := FALSE,
       RequestedContactor1 := FALSE, RequestedContactor2 := FALSE,
       RequestedContactor3 := FALSE, RequestedContactor4 := FALSE,
       RequestedStep := 0, DropConfirmDelay := T#300ms, MaxSenseHoldTime := T#1s);
    ADVANCE_TIME(10000000);
fb(Enable := TRUE, Reset := FALSE, SafeStop := FALSE, AscentPermit := TRUE, DescendPermit := TRUE, PowerContactorEngaged := TRUE,
       BrakeFeedback := TRUE, FwdRevSpeedFeedbackOff := TRUE,
       RequestedRelayFwd := TRUE, RequestedRelayRev := FALSE,
       RequestedContactor1 := FALSE, RequestedContactor2 := FALSE,
       RequestedContactor3 := FALSE, RequestedContactor4 := FALSE,
       RequestedStep := 0, DropConfirmDelay := T#300ms, MaxSenseHoldTime := T#1s);
    ASSERT_FALSE(fb.RelayFwd, 'Confirmation retombee -> chute du sens (§3bis)');
    ASSERT_FALSE(fb.BrakeCmd, 'Apres chute -> BrakeCmd=FALSE');
    ASSERT_FALSE(fb.SenseHoldActive, 'Fin du maintien');
    ASSERT_EQ(fb.State, E_WinchFinalInterlockState.READY, 'Retour READY');
END_TEST

TEST 'TC-P10-023b §3bis : T_max atteint sans confirmation -> chute du sens FORCEE + latch ContactorStuck'
    (* FwdRevSpeedFeedbackOff reste FALSE (contacteurs ne confirment pas la retombee). Apres
       MaxSenseHoldTime (T_max=300ms) la barriere FORCE la chute du sens et latche
       ContactorStuck (AC7). Le maintien indefini du stator est interdit. *)
    fb(Enable := TRUE, Reset := FALSE, SafeStop := FALSE, AscentPermit := TRUE, DescendPermit := TRUE, PowerContactorEngaged := TRUE,
       BrakeFeedback := FALSE, FwdRevSpeedFeedbackOff := TRUE,
       RequestedRelayFwd := FALSE, RequestedRelayRev := FALSE,
       RequestedContactor1 := FALSE, RequestedContactor2 := FALSE,
       RequestedContactor3 := FALSE, RequestedContactor4 := FALSE,
       RequestedStep := 0, DropConfirmDelay := T#200ms, MaxSenseHoldTime := T#300ms);
    ADVANCE_TIME(1500000000);
fb(Enable := TRUE, Reset := FALSE, SafeStop := FALSE, AscentPermit := TRUE, DescendPermit := TRUE, PowerContactorEngaged := TRUE,
       BrakeFeedback := FALSE, FwdRevSpeedFeedbackOff := TRUE,
       RequestedRelayFwd := FALSE, RequestedRelayRev := FALSE,
       RequestedContactor1 := FALSE, RequestedContactor2 := FALSE,
       RequestedContactor3 := FALSE, RequestedContactor4 := FALSE,
       RequestedStep := 0, DropConfirmDelay := T#200ms, MaxSenseHoldTime := T#300ms);

    (* Scan 2 : mouvement montee *)
    ADVANCE_TIME(10000000);
fb(Enable := TRUE, Reset := FALSE, SafeStop := FALSE, AscentPermit := TRUE, DescendPermit := TRUE, PowerContactorEngaged := TRUE,
       BrakeFeedback := TRUE, FwdRevSpeedFeedbackOff := FALSE,
       RequestedRelayFwd := TRUE, RequestedRelayRev := FALSE,
       RequestedContactor1 := TRUE, RequestedContactor2 := FALSE,
       RequestedContactor3 := FALSE, RequestedContactor4 := FALSE,
       RequestedStep := 1, DropConfirmDelay := T#200ms, MaxSenseHoldTime := T#300ms);
    ASSERT_TRUE(fb.RelayFwd, 'Mouvement -> RelayFwd');

    (* Scan 3 : chute palier a 0, sens maintenu, MAIS contacteurs jamais confirmes retombes *)
    ADVANCE_TIME(10000000);
fb(Enable := TRUE, Reset := FALSE, SafeStop := FALSE, AscentPermit := TRUE, DescendPermit := TRUE, PowerContactorEngaged := TRUE,
       BrakeFeedback := TRUE, FwdRevSpeedFeedbackOff := FALSE,
       RequestedRelayFwd := TRUE, RequestedRelayRev := FALSE,
       RequestedContactor1 := FALSE, RequestedContactor2 := FALSE,
       RequestedContactor3 := FALSE, RequestedContactor4 := FALSE,
       RequestedStep := 0, DropConfirmDelay := T#200ms, MaxSenseHoldTime := T#300ms);
    ASSERT_TRUE(fb.RelayFwd, 'Entree en maintien -> sens tenu');
    ASSERT_TRUE(fb.SenseHoldActive, 'SenseHoldActive');

    (* Scan 4 : T_max (300ms) depasse sans confirmation -> chute forcee + latch *)
    ADVANCE_TIME(10000000);
fb(Enable := TRUE, Reset := FALSE, SafeStop := FALSE, AscentPermit := TRUE, DescendPermit := TRUE, PowerContactorEngaged := TRUE,
       BrakeFeedback := TRUE, FwdRevSpeedFeedbackOff := FALSE,
       RequestedRelayFwd := TRUE, RequestedRelayRev := FALSE,
       RequestedContactor1 := FALSE, RequestedContactor2 := FALSE,
       RequestedContactor3 := FALSE, RequestedContactor4 := FALSE,
       RequestedStep := 0, DropConfirmDelay := T#200ms, MaxSenseHoldTime := T#300ms);
    ADVANCE_TIME(400000000);
fb(Enable := TRUE, Reset := FALSE, SafeStop := FALSE, AscentPermit := TRUE, DescendPermit := TRUE, PowerContactorEngaged := TRUE,
       BrakeFeedback := TRUE, FwdRevSpeedFeedbackOff := FALSE,
       RequestedRelayFwd := TRUE, RequestedRelayRev := FALSE,
       RequestedContactor1 := FALSE, RequestedContactor2 := FALSE,
       RequestedContactor3 := FALSE, RequestedContactor4 := FALSE,
       RequestedStep := 0, DropConfirmDelay := T#200ms, MaxSenseHoldTime := T#300ms);
    ASSERT_FALSE(fb.RelayFwd, 'T_max sans confirmation -> chute du sens FORCEE (AC7)');
    ASSERT_FALSE(fb.BrakeCmd, 'Chute forcee -> BrakeCmd=FALSE');
    ASSERT_TRUE(fb.ContactorStuck, 'Diag ContactorStuck latche');
    ASSERT_FALSE(fb.SenseHoldActive, 'Fin du maintien');
    ASSERT_FALSE(fb.Ready, 'Latch -> barriere non pret (pas de redemarrage auto)');
    ASSERT_EQ(fb.State, E_WinchFinalInterlockState.FAULT, 'Etat FAULT');
    ASSERT_EQ(fb.Reason, E_WinchFinalInterlockReason.SENSE_DROP_TIMEOUT, 'Reason=SENSE_DROP_TIMEOUT');

    (* Scan 5 : acquittement conscient (front Reset) -> latch leve (cause disparue = demande neutre) *)
    ADVANCE_TIME(10000000);
    fb(Enable := TRUE, Reset := TRUE, SafeStop := FALSE, PowerContactorEngaged := TRUE,
       BrakeFeedback := TRUE, FwdRevSpeedFeedbackOff := TRUE,
       RequestedRelayFwd := FALSE, RequestedRelayRev := FALSE,
       RequestedContactor1 := FALSE, RequestedContactor2 := FALSE,
       RequestedContactor3 := FALSE, RequestedContactor4 := FALSE,
       RequestedStep := 0, DropConfirmDelay := T#200ms, MaxSenseHoldTime := T#300ms);
    ADVANCE_TIME(10000000);
fb(Enable := TRUE, Reset := FALSE, SafeStop := FALSE, AscentPermit := TRUE, DescendPermit := TRUE, PowerContactorEngaged := TRUE,
       BrakeFeedback := TRUE, FwdRevSpeedFeedbackOff := TRUE,
       RequestedRelayFwd := FALSE, RequestedRelayRev := FALSE,
       RequestedContactor1 := FALSE, RequestedContactor2 := FALSE,
       RequestedContactor3 := FALSE, RequestedContactor4 := FALSE,
       RequestedStep := 0, DropConfirmDelay := T#200ms, MaxSenseHoldTime := T#300ms);
    ASSERT_FALSE(fb.ContactorStuck, 'Front Reset conscient -> latch ContactorStuck leve');
END_TEST

TEST 'TC-P10-023c §3bis : coupure dure (Enable=FALSE) pendant le maintien -> RelayFwd=FALSE immediat'
    (* La coupure dure ne passe JAMAIS par le maintien §3bis (AC9) : Enable=FALSE en pleine
       tenue du sens coupe RelayFwd/Rev au cycle suivant, sans attendre confirmation ni T_max. *)
    fb(Enable := TRUE, Reset := FALSE, SafeStop := FALSE, AscentPermit := TRUE, DescendPermit := TRUE, PowerContactorEngaged := TRUE,
       BrakeFeedback := FALSE, FwdRevSpeedFeedbackOff := TRUE,
       RequestedRelayFwd := FALSE, RequestedRelayRev := FALSE,
       RequestedContactor1 := FALSE, RequestedContactor2 := FALSE,
       RequestedContactor3 := FALSE, RequestedContactor4 := FALSE,
       RequestedStep := 0, DropConfirmDelay := T#300ms, MaxSenseHoldTime := T#1s);
    ADVANCE_TIME(1500000000);
fb(Enable := TRUE, Reset := FALSE, SafeStop := FALSE, AscentPermit := TRUE, DescendPermit := TRUE, PowerContactorEngaged := TRUE,
       BrakeFeedback := FALSE, FwdRevSpeedFeedbackOff := TRUE,
       RequestedRelayFwd := FALSE, RequestedRelayRev := FALSE,
       RequestedContactor1 := FALSE, RequestedContactor2 := FALSE,
       RequestedContactor3 := FALSE, RequestedContactor4 := FALSE,
       RequestedStep := 0, DropConfirmDelay := T#300ms, MaxSenseHoldTime := T#1s);

    (* Scan 2 : mouvement montee *)
    ADVANCE_TIME(10000000);
fb(Enable := TRUE, Reset := FALSE, SafeStop := FALSE, AscentPermit := TRUE, DescendPermit := TRUE, PowerContactorEngaged := TRUE,
       BrakeFeedback := TRUE, FwdRevSpeedFeedbackOff := FALSE,
       RequestedRelayFwd := TRUE, RequestedRelayRev := FALSE,
       RequestedContactor1 := TRUE, RequestedContactor2 := FALSE,
       RequestedContactor3 := FALSE, RequestedContactor4 := FALSE,
       RequestedStep := 1, DropConfirmDelay := T#300ms, MaxSenseHoldTime := T#1s);
    ASSERT_TRUE(fb.RelayFwd, 'Mouvement -> RelayFwd');

    (* Scan 3 : chute palier a 0 -> maintien actif *)
    ADVANCE_TIME(10000000);
fb(Enable := TRUE, Reset := FALSE, SafeStop := FALSE, AscentPermit := TRUE, DescendPermit := TRUE, PowerContactorEngaged := TRUE,
       BrakeFeedback := TRUE, FwdRevSpeedFeedbackOff := FALSE,
       RequestedRelayFwd := TRUE, RequestedRelayRev := FALSE,
       RequestedContactor1 := FALSE, RequestedContactor2 := FALSE,
       RequestedContactor3 := FALSE, RequestedContactor4 := FALSE,
       RequestedStep := 0, DropConfirmDelay := T#300ms, MaxSenseHoldTime := T#1s);
    ASSERT_TRUE(fb.RelayFwd, 'Maintien actif -> sens tenu');
    ASSERT_TRUE(fb.SenseHoldActive, 'SenseHoldActive');

    (* Scan 4 : Enable=FALSE -> coupure dure immediate, meme en pleine tenue *)
    ADVANCE_TIME(10000000);
    fb(Enable := FALSE, Reset := FALSE, SafeStop := FALSE, PowerContactorEngaged := TRUE,
       BrakeFeedback := TRUE, FwdRevSpeedFeedbackOff := FALSE,
       RequestedRelayFwd := TRUE, RequestedRelayRev := FALSE,
       RequestedContactor1 := FALSE, RequestedContactor2 := FALSE,
       RequestedContactor3 := FALSE, RequestedContactor4 := FALSE,
       RequestedStep := 0, DropConfirmDelay := T#300ms, MaxSenseHoldTime := T#1s);
    ASSERT_FALSE(fb.RelayFwd, 'Enable=FALSE -> RelayFwd=FALSE immediat (AC9)');
    ASSERT_FALSE(fb.BrakeCmd, 'Enable=FALSE -> BrakeCmd=FALSE immediat');
    ASSERT_FALSE(fb.SenseHoldActive, 'Maintien neutralise par la gate');
END_TEST

TEST 'TC-T216-FINAL-PERMIT Direction refusee coupe la barriere finale, direction autorisee passe'
    (* Le permis final est une defense en profondeur : il doit couper relais,
       contacteurs et frein meme si une demande physique est encore presente. *)
    fb(Enable := TRUE, Reset := FALSE, SafeStop := FALSE, AscentPermit := TRUE, DescendPermit := TRUE,
       PowerContactorEngaged := TRUE, BrakeFeedback := TRUE, FwdRevSpeedFeedbackOff := TRUE,
       RequestedRelayFwd := TRUE, RequestedRelayRev := FALSE,
       RequestedContactor1 := TRUE, RequestedContactor2 := FALSE,
       RequestedContactor3 := FALSE, RequestedContactor4 := FALSE, RequestedStep := 1);
    ASSERT_TRUE(fb.RelayFwd, 'Permis montee TRUE -> relais montee autorise');
    ASSERT_TRUE(fb.BrakeCmd, 'Permis montee TRUE -> frein desserre');

    ADVANCE_TIME(10000000);
    fb(Enable := TRUE, Reset := FALSE, SafeStop := FALSE, AscentPermit := FALSE, DescendPermit := TRUE,
       PowerContactorEngaged := TRUE, BrakeFeedback := TRUE, FwdRevSpeedFeedbackOff := TRUE,
       RequestedRelayFwd := TRUE, RequestedRelayRev := FALSE,
       RequestedContactor1 := TRUE, RequestedContactor2 := FALSE,
       RequestedContactor3 := FALSE, RequestedContactor4 := FALSE, RequestedStep := 1);
    ASSERT_FALSE(fb.RelayFwd, 'Permis montee FALSE -> relais montee coupe');
    ASSERT_FALSE(fb.Contactor1, 'Permis montee FALSE -> contacteur coupe');
    ASSERT_FALSE(fb.BrakeCmd, 'Permis montee FALSE -> frein serre');

    ADVANCE_TIME(10000000);
    fb(Enable := TRUE, Reset := FALSE, SafeStop := FALSE, AscentPermit := TRUE, DescendPermit := FALSE,
       PowerContactorEngaged := TRUE, BrakeFeedback := TRUE, FwdRevSpeedFeedbackOff := TRUE,
       RequestedRelayFwd := FALSE, RequestedRelayRev := TRUE,
       RequestedContactor1 := TRUE, RequestedContactor2 := FALSE,
       RequestedContactor3 := FALSE, RequestedContactor4 := FALSE, RequestedStep := 1);
    ASSERT_FALSE(fb.RelayRev, 'Permis descente FALSE -> relais descente coupe');
    ASSERT_FALSE(fb.Contactor1, 'Permis descente FALSE -> contacteur coupe');
    ASSERT_FALSE(fb.BrakeCmd, 'Permis descente FALSE -> frein serre');
END_TEST

(* ---- test_fb_winchstepshaper.st ---- *)
SETUP
VAR
    fb : FB_WinchStepShaper;
END_VAR
END_SETUP

TEST 'TC-P10-SHAPER-01 Montee nominale 1000ms'
    fb(Enable := TRUE, TargetStep := 0, StepRampDelay := T#1000ms);
    ASSERT_EQ(fb.ShapedStep, 0, 'ShapedStep initialement a 0');

    (* Depart immediat 0->1 au scan 0 *)
    fb(Enable := TRUE, TargetStep := 5, StepRampDelay := T#1000ms);
    ASSERT_EQ(fb.ShapedStep, 1, 'ShapedStep passe a 1 immediatement');

    (* Echantillonnage avant delai *)
    ADVANCE_TIME(10000000);
    fb(Enable := TRUE, TargetStep := 5, StepRampDelay := T#1000ms);
    ASSERT_EQ(fb.ShapedStep, 1, 'Reste a 1 avant delai');

    (* Ecoulement 1000ms -> P2 *)
    ADVANCE_TIME(1000000000);
    fb(Enable := TRUE, TargetStep := 5, StepRampDelay := T#1000ms);
    ASSERT_EQ(fb.ShapedStep, 2, 'Passe a 2 apres delai');
END_TEST

TEST 'TC-P10-SHAPER-02 Descente nominale 500ms'
    fb(Enable := TRUE, TargetStep := 2, StepRampDelay := T#500ms);
    ASSERT_EQ(fb.ShapedStep, 1, 'Depart P1');

    ADVANCE_TIME(10000000);
    fb(Enable := TRUE, TargetStep := 2, StepRampDelay := T#500ms);
    ASSERT_EQ(fb.ShapedStep, 1, 'Reste a 1');

    ADVANCE_TIME(500000000);
    fb(Enable := TRUE, TargetStep := 2, StepRampDelay := T#500ms);
    ASSERT_EQ(fb.ShapedStep, 2, 'Passe a 2 apres delai 500ms');
END_TEST

TEST 'TC-P10-SHAPER-03 Asymetrie arret direct'
    fb(Enable := TRUE, TargetStep := 2, StepRampDelay := T#500ms);
    ASSERT_EQ(fb.ShapedStep, 1, 'Depart P1');

    ADVANCE_TIME(10000000);
    fb(Enable := TRUE, TargetStep := 2, StepRampDelay := T#500ms);
    ADVANCE_TIME(500000000);
    fb(Enable := TRUE, TargetStep := 2, StepRampDelay := T#500ms);
    ASSERT_EQ(fb.ShapedStep, 2, 'P2 etabli');

    (* Descente a 1 immediate *)
    fb(Enable := TRUE, TargetStep := 1, StepRampDelay := T#500ms);
    ASSERT_EQ(fb.ShapedStep, 1, 'Descente immediate a la cible P1');

    (* Arret franc *)
    fb(Enable := TRUE, TargetStep := 0, StepRampDelay := T#500ms);
    ASSERT_EQ(fb.ShapedStep, 0, 'Arret immediat a 0');
END_TEST

TEST 'TC-P10-SHAPER-04 Rejet hors plage'
    fb(Enable := TRUE, TargetStep := 2, StepRampDelay := T#500ms);
    ASSERT_EQ(fb.ShapedStep, 1, 'Depart P1');

    fb(Enable := FALSE, TargetStep := 2, StepRampDelay := T#500ms);
    ASSERT_EQ(fb.ShapedStep, 0, 'Enable FALSE remet a 0');
END_TEST

(* ---- test_fb_winchsync.st ---- *)
(* =======================================================================
   🧪 test_fb_winchsync.st — FB_WinchSync (TC-P10-014, 015, 016)
   ───────────────────────────────────────────────────────────────
   Fiche : DOC/AF/AF_Partie-10_Fonction_Winch/FB_WinchSync_v1.1.md
   Conventions : 1 appel fb() = 1 scan ; ADVANCE_TIME(10000000) entre les
   scans pour les fronts R_TRIG.
   Seuils (v1.1) : Warn = CfgSyncToleranceM=0.8m (instantané + latch, sans timer) ;
   Fault = CfgSyncCriticalToleranceM=0.50m (filtre 800ms) ; incohérence commande = 500ms.
   ======================================================================= *)

SETUP
VAR
    fb : FB_WinchSync;
END_VAR
END_SETUP

(* ── Remise à zéro commune : Enable=TRUE, Mode MAINT_N1 (SyncActive imposé), positions alignées ── *)

TEST 'TC-P10-014 Ecart M1/M2 > seuil Warn (0.8m) : SyncWarn instantane + latch, sans timer, pas de coupure'
    (* Scan 1 : regime nominal, positions alignees *)
    fb(Enable := TRUE, Reset := FALSE, Mode := E_Mode.MAINT_N1, SyncEnable := TRUE,
       CablePosM1 := 0.0, CablePosM2 := 0.0,
       HomedAndReliableM1 := TRUE, HomedAndReliableM2 := TRUE,
       CfgSyncToleranceM := 0.8, CfgSyncCriticalToleranceM := 0.50, ActiveOffsetM := 0.0);
    ADVANCE_TIME(10000000);
    fb(Enable := TRUE, Reset := FALSE, Mode := E_Mode.MAINT_N1, SyncEnable := TRUE,
       CablePosM1 := 0.0, CablePosM2 := 0.0,
       HomedAndReliableM1 := TRUE, HomedAndReliableM2 := TRUE,
       CfgSyncToleranceM := 0.8, CfgSyncCriticalToleranceM := 0.50, ActiveOffsetM := 0.0);
    ASSERT_TRUE(fb.SyncActive, 'Mode MAINT_N1 -> SyncActive=TRUE');
    ASSERT_FALSE(fb.SyncDeviationWarn, 'Positions alignees -> pas de Warn');

    (* Scan 2 : ecart M1/M2 = 1.0m > 0.8m -> Warn instantane (sans timer) *)
    ADVANCE_TIME(10000000);
    fb(Enable := TRUE, Reset := FALSE, Mode := E_Mode.MAINT_N1, SyncEnable := TRUE,
       CablePosM1 := 1.0, CablePosM2 := 0.0,
       HomedAndReliableM1 := TRUE, HomedAndReliableM2 := TRUE,
       CfgSyncToleranceM := 0.8, CfgSyncCriticalToleranceM := 0.50, ActiveOffsetM := 0.0);
    ASSERT_TRUE(fb.SyncDeviationWarn, 'Ecart >0.8m -> SyncDeviationWarn instantane');
    ASSERT_TRUE(fb.SyncWarn, 'Ecart >0.8m -> SyncWarn IHM');
    ASSERT_TRUE(fb.Fault.Error, 'Ecart >0.8m -> Error');

    (* Scan 3 : cause disparue -> Warn LATCHE (reste actif sans timer) *)
    ADVANCE_TIME(10000000);
    fb(Enable := TRUE, Reset := FALSE, Mode := E_Mode.MAINT_N1, SyncEnable := TRUE,
       CablePosM1 := 0.0, CablePosM2 := 0.0,
       HomedAndReliableM1 := TRUE, HomedAndReliableM2 := TRUE,
       CfgSyncToleranceM := 0.8, CfgSyncCriticalToleranceM := 0.50, ActiveOffsetM := 0.0);
    ASSERT_TRUE(fb.SyncDeviationWarn, 'Cause disparue -> Warn latche conserve');

    (* Scan 4 : front Reset -> Warn leve *)
    ADVANCE_TIME(10000000);
    fb(Enable := TRUE, Reset := TRUE, Mode := E_Mode.MAINT_N1, SyncEnable := TRUE,
       CablePosM1 := 0.0, CablePosM2 := 0.0,
       HomedAndReliableM1 := TRUE, HomedAndReliableM2 := TRUE,
       CfgSyncToleranceM := 0.8, CfgSyncCriticalToleranceM := 0.50, ActiveOffsetM := 0.0);
    ADVANCE_TIME(10000000);
    fb(Enable := TRUE, Reset := FALSE, Mode := E_Mode.MAINT_N1, SyncEnable := TRUE,
       CablePosM1 := 0.0, CablePosM2 := 0.0,
       HomedAndReliableM1 := TRUE, HomedAndReliableM2 := TRUE,
       CfgSyncToleranceM := 0.8, CfgSyncCriticalToleranceM := 0.50, ActiveOffsetM := 0.0);
    ASSERT_FALSE(fb.SyncDeviationWarn, 'Reset -> Warn leve');
    ASSERT_FALSE(fb.SyncWarn, 'Reset -> SyncWarn leve');
END_TEST

TEST 'T258-REX-20260906 Gate ferme purge le warning deviation avant reactivation'
    (* Reproduit la trace terrain : un ecart avertissement est memorise avant
       une phase dissymetrique, puis le gate est coupe et reactive avec 0.088 m. *)
    fb(Enable := TRUE, Reset := FALSE, Mode := E_Mode.SEMI_AUTO, SyncEnable := TRUE,
       CablePosM1 := -3.210, CablePosM2 := 0.0,
       HomedAndReliableM1 := TRUE, HomedAndReliableM2 := TRUE,
       CfgSyncToleranceM := 3.0, CfgSyncCriticalToleranceM := 6.0, ActiveOffsetM := 0.0);
    ASSERT_TRUE(fb.SyncDeviationWarn, 'Ecart 3.210m > seuil 3m : warning memorise');

    ADVANCE_TIME(10000000);
    fb(Enable := FALSE, Reset := FALSE);
    ASSERT_FALSE(fb.Fault.Error, 'Gate ferme : aucun defaut publie');

    ADVANCE_TIME(10000000);
    fb(Enable := TRUE, Reset := FALSE, Mode := E_Mode.SEMI_AUTO, SyncEnable := TRUE,
       CablePosM1 := 0.088, CablePosM2 := 0.0,
       HomedAndReliableM1 := TRUE, HomedAndReliableM2 := TRUE,
       CfgSyncToleranceM := 3.0, CfgSyncCriticalToleranceM := 6.0, ActiveOffsetM := 0.0);
    ASSERT_FALSE(fb.SyncDeviationWarn, 'Reactivation sous seuil : aucun warning residuel');
    ASSERT_FALSE(fb.Fault.Error, 'Reactivation sous seuil : Error reste FALSE');
    ASSERT_EQ(fb.Fault.ErrorId, 0, 'Reactivation sous seuil : ErrorId remis a zero');
END_TEST

TEST 'TC-P10-014bis Ecart > seuil Fault (0.50m) : SyncDeviationFault filtre 800ms'
    (* Scan 1 : regime nominal *)
    fb(Enable := TRUE, Reset := FALSE, Mode := E_Mode.MAINT_N1, SyncEnable := TRUE,
       CablePosM1 := 0.0, CablePosM2 := 0.0,
       HomedAndReliableM1 := TRUE, HomedAndReliableM2 := TRUE,
       CfgSyncToleranceM := 0.8, CfgSyncCriticalToleranceM := 0.50, ActiveOffsetM := 0.0);
    ADVANCE_TIME(10000000);
    fb(Enable := TRUE, Reset := FALSE, Mode := E_Mode.MAINT_N1, SyncEnable := TRUE,
       CablePosM1 := 0.0, CablePosM2 := 0.0,
       HomedAndReliableM1 := TRUE, HomedAndReliableM2 := TRUE,
       CfgSyncToleranceM := 0.8, CfgSyncCriticalToleranceM := 0.50, ActiveOffsetM := 0.0);

    (* Scan 2 : ecart = 1.0m > 0.50m -> Fault filtre 800ms (pas immediat) *)
    ADVANCE_TIME(10000000);
    fb(Enable := TRUE, Reset := FALSE, Mode := E_Mode.MAINT_N1, SyncEnable := TRUE,
       CablePosM1 := 1.0, CablePosM2 := 0.0,
       HomedAndReliableM1 := TRUE, HomedAndReliableM2 := TRUE,
       CfgSyncToleranceM := 0.8, CfgSyncCriticalToleranceM := 0.50, ActiveOffsetM := 0.0);
    ASSERT_FALSE(fb.SyncDeviationFault, 'Avant 800ms : pas de Fault (filtre transitoire)');

    (* Scan 3 : apres 800ms -> SyncDeviationFault *)
    ADVANCE_TIME(800000000);
    fb(Enable := TRUE, Reset := FALSE, Mode := E_Mode.MAINT_N1, SyncEnable := TRUE,
       CablePosM1 := 1.0, CablePosM2 := 0.0,
       HomedAndReliableM1 := TRUE, HomedAndReliableM2 := TRUE,
       CfgSyncToleranceM := 0.8, CfgSyncCriticalToleranceM := 0.50, ActiveOffsetM := 0.0);
    ASSERT_TRUE(fb.SyncDeviationFault, 'Ecart >0.50m 800ms -> SyncDeviationFault');
    ASSERT_TRUE(fb.SyncWarn, 'Fault -> SyncWarn');
END_TEST

TEST 'TC-P10-015 Incoherence commande (bit1) : discordance contacteurs 500ms -> SyncWarn'
    (* Scan 1 : regime nominal, commandes identiques *)
    fb(Enable := TRUE, Reset := FALSE, Mode := E_Mode.MAINT_N1, SyncEnable := TRUE,
       CablePosM1 := 0.0, CablePosM2 := 0.0,
       HomedAndReliableM1 := TRUE, HomedAndReliableM2 := TRUE,
       CfgSyncToleranceM := 0.8, CfgSyncCriticalToleranceM := 0.50, ActiveOffsetM := 0.0,
       RelayFwdM1 := TRUE, RelayFwdM2 := TRUE,
       RelayRevM1 := FALSE, RelayRevM2 := FALSE,
       Contactor1_M1 := TRUE, Contactor1_M2 := TRUE,
       Contactor2_M1 := FALSE, Contactor2_M2 := FALSE,
       Contactor3_M1 := FALSE, Contactor3_M2 := FALSE,
       Contactor4_M1 := FALSE, Contactor4_M2 := FALSE);
    ADVANCE_TIME(10000000);
    fb(Enable := TRUE, Reset := FALSE, Mode := E_Mode.MAINT_N1, SyncEnable := TRUE,
       CablePosM1 := 0.0, CablePosM2 := 0.0,
       HomedAndReliableM1 := TRUE, HomedAndReliableM2 := TRUE,
       CfgSyncToleranceM := 0.8, CfgSyncCriticalToleranceM := 0.50, ActiveOffsetM := 0.0,
       RelayFwdM1 := TRUE, RelayFwdM2 := TRUE,
       RelayRevM1 := FALSE, RelayRevM2 := FALSE,
       Contactor1_M1 := TRUE, Contactor1_M2 := TRUE,
       Contactor2_M1 := FALSE, Contactor2_M2 := FALSE,
       Contactor3_M1 := FALSE, Contactor3_M2 := FALSE,
       Contactor4_M1 := FALSE, Contactor4_M2 := FALSE);
    ASSERT_FALSE(fb.SyncWarn, 'Commandes identiques -> pas de Warn');

    (* Scan 2 : discordance RelayFwdM1=TRUE vs RelayFwdM2=FALSE -> filtre 500ms *)
    ADVANCE_TIME(10000000);
    fb(Enable := TRUE, Reset := FALSE, Mode := E_Mode.MAINT_N1, SyncEnable := TRUE,
       CablePosM1 := 0.0, CablePosM2 := 0.0,
       HomedAndReliableM1 := TRUE, HomedAndReliableM2 := TRUE,
       CfgSyncToleranceM := 0.8, CfgSyncCriticalToleranceM := 0.50, ActiveOffsetM := 0.0,
       RelayFwdM1 := TRUE, RelayFwdM2 := FALSE,
       RelayRevM1 := FALSE, RelayRevM2 := FALSE,
       Contactor1_M1 := TRUE, Contactor1_M2 := TRUE,
       Contactor2_M1 := FALSE, Contactor2_M2 := FALSE,
       Contactor3_M1 := FALSE, Contactor3_M2 := FALSE,
       Contactor4_M1 := FALSE, Contactor4_M2 := FALSE);
    ASSERT_FALSE(fb.SyncWarn, 'Avant 500ms : pas encore de Warn (filtre)');

    (* Scan 3 : apres 500ms -> ContactorMismatch -> SyncWarn *)
    ADVANCE_TIME(500000000);
    fb(Enable := TRUE, Reset := FALSE, Mode := E_Mode.MAINT_N1, SyncEnable := TRUE,
       CablePosM1 := 0.0, CablePosM2 := 0.0,
       HomedAndReliableM1 := TRUE, HomedAndReliableM2 := TRUE,
       CfgSyncToleranceM := 0.8, CfgSyncCriticalToleranceM := 0.50, ActiveOffsetM := 0.0,
       RelayFwdM1 := TRUE, RelayFwdM2 := FALSE,
       RelayRevM1 := FALSE, RelayRevM2 := FALSE,
       Contactor1_M1 := TRUE, Contactor1_M2 := TRUE,
       Contactor2_M1 := FALSE, Contactor2_M2 := FALSE,
       Contactor3_M1 := FALSE, Contactor3_M2 := FALSE,
       Contactor4_M1 := FALSE, Contactor4_M2 := FALSE);
    ASSERT_TRUE(fb.SyncWarn, 'Discordance contacteurs 500ms -> SyncWarn');
    ASSERT_TRUE(fb.Fault.Error, 'Discordance -> Error');
END_TEST

TEST 'TC-P10-016 Couplage croise : SyncActive=TRUE conditionne la coupure M2 au meme scan'
    (* (essai site — stub) : la coupure croisee reelle (SafeStopM2_Active := SafeStopM2_Raw OR
       (SyncActive AND SafeStopM1_Raw)) est cablee dans PRG_04_Treuils_Benne.st, pas dans ce FB.
       On verifie ici la brique amont : SyncActive=TRUE (condition du couplage) selon le mode. *)
    (* Mode MAINT_N1 -> SyncActive impose TRUE *)
    fb(Enable := TRUE, Reset := FALSE, Mode := E_Mode.MAINT_N1, SyncEnable := FALSE,
       CablePosM1 := 0.0, CablePosM2 := 0.0,
       HomedAndReliableM1 := TRUE, HomedAndReliableM2 := TRUE,
       CfgSyncToleranceM := 0.8, CfgSyncCriticalToleranceM := 0.50, ActiveOffsetM := 0.0);
    ASSERT_TRUE(fb.SyncActive, 'MAINT_N1 -> SyncActive=TRUE (couplage actif)');

    (* Mode MAINT_N2 -> SyncActive = SyncEnable (pilotable) *)
    ADVANCE_TIME(10000000);
    fb(Enable := TRUE, Reset := FALSE, Mode := E_Mode.MAINT_N2, SyncEnable := FALSE,
       CablePosM1 := 0.0, CablePosM2 := 0.0,
       HomedAndReliableM1 := TRUE, HomedAndReliableM2 := TRUE,
       CfgSyncToleranceM := 0.8, CfgSyncCriticalToleranceM := 0.50, ActiveOffsetM := 0.0);
    ASSERT_FALSE(fb.SyncActive, 'MAINT_N2 + SyncEnable=FALSE -> SyncActive=FALSE');
    ADVANCE_TIME(10000000);
    fb(Enable := TRUE, Reset := FALSE, Mode := E_Mode.MAINT_N2, SyncEnable := TRUE,
       CablePosM1 := 0.0, CablePosM2 := 0.0,
       HomedAndReliableM1 := TRUE, HomedAndReliableM2 := TRUE,
       CfgSyncToleranceM := 0.8, CfgSyncCriticalToleranceM := 0.50, ActiveOffsetM := 0.0);
    ASSERT_TRUE(fb.SyncActive, 'MAINT_N2 + SyncEnable=TRUE -> SyncActive=TRUE');
END_TEST
